Fanuc KAREL source: kb00010.KL

-- PROVISIONAL review KL for V770-1; original PC SHA256 87165fae012a7bf2b04327fd018944051831a459ccf05e4026ff639894b07331
-- Incomplete behavior may be omitted. Consult companion uncertainty JSON. Do not deploy.
PROGRAM KB00010
%NOLOCKGROUP
BEGIN
  -- UNRESOLVED_PC offsets 5-14; opcodes 3F,75
  -- UNRESOLVED_PC offsets 19-28; opcodes 3F,75
  -- UNRESOLVED_PC offsets 33-40; opcodes 9D,23
  -- UNRESOLVED_PC offsets 45-52; opcodes 9D,23
  -- UNRESOLVED_PC offsets 57-66; opcodes 3F,75
  -- UNRESOLVED_PC offsets 71-78; opcodes 9D,23
  -- UNRESOLVED_PC offsets 83-129; opcodes 27,22,2A,22,2A,22,22,22,2A,22,31
  -- UNRESOLVED_PC offsets 134-138; opcodes 7F
END KB00010
